(* IEC 61131-3 sources: laba_2_/Libraries/DriveLib, 3 files *)

(* ---- Types.typ ---- *)
TYPE
	states_door :
		(
		ST_INIT := 1,
		ST_UNKNOWN := 2,
		ST_OPEN := 3,
		ST_CLOSE := 4,
		ST_ACC_POS := 5,
		ST_ACC_NEG := 6,
		ST_POS := 7,
		ST_NEG := 8,
		ST_DEC_POS := 9,
		ST_DEC_NEG := 10
		);
END_TYPE

(* ---- Constants.var ---- *)
VAR CONSTANT
	CMD_ENABLE : USINT := 15;
	CMD_SWITCH_ON : USINT := 7;
	CMD_SHUTDOWN : USINT := 6;
	STATE_DISABLED : USINT := 64;
	STATE_SWITCHED_ON : USINT := 35;
	STATE_READY : USINT := 33;
END_VAR

(* ---- DriveLib.fun ---- *)
{REDUND_ERROR} FUNCTION_BLOCK DriveStateMashine (*TODO: Add your comment here*) (*$GROUP=User,$CAT=User,$GROUPICON=User.png,$CATICON=User.png*)
	VAR_INPUT
		state : {REDUND_UNREPLICABLE} UINT;
		enable : BOOL;
	END_VAR
	VAR_OUTPUT
		command : UINT;
		speed : INT;
	END_VAR
END_FUNCTION_BLOCK

{REDUND_ERROR} FUNCTION_BLOCK DoorStateMashine (*TODO: Add your comment here*) (*$GROUP=User,$CAT=User,$GROUPICON=User.png,$CATICON=User.png*)
	VAR_INPUT
		state : UINT;
		sw1 : BOOL;
		sw2 : BOOL;
		sw3 : BOOL;
		sw4 : BOOL;
		direction : BOOL;
	END_VAR
	VAR_OUTPUT
		speed : INT;
	END_VAR
END_FUNCTION_BLOCK

{REDUND_ERROR} {REDUND_UNREPLICABLE} FUNCTION_BLOCK LedStateMashine (*TODO: Add your comment here*) (*$GROUP=User,$CAT=User,$GROUPICON=User.png,$CATICON=User.png*)
	VAR_INPUT
		state : {REDUND_UNREPLICABLE} UINT;
	END_VAR
	VAR_OUTPUT
		led1 : {REDUND_UNREPLICABLE} BOOL;
		led2 : {REDUND_UNREPLICABLE} BOOL;
		led3 : {REDUND_UNREPLICABLE} BOOL;
		led4 : {REDUND_UNREPLICABLE} BOOL;
		timer : {REDUND_UNREPLICABLE} INT;
	END_VAR
END_FUNCTION_BLOCK
